FUNCTION_BLOCK ReactorAbortManager (* Basic Function Block Type *)
  (* Standard: 61499-2 *)
  (* Version 0.0, 10/19/2026, Schneider Electric, Template *)
  PACKAGE SE.Nereda;
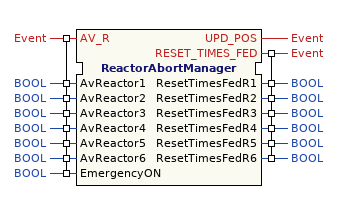
  EVENT_INPUT
    AV_R WITH AvReactor1, AvReactor2, AvReactor3, AvReactor4, AvReactor5, AvReactor6, EmergencyON; (* Normal Execution Request *)
  END_EVENT
  EVENT_OUTPUT
    UPD_POS; (* Execution Confirmation *)
    RESET_TIMES_FED WITH ResetTimesFedR1, ResetTimesFedR2, ResetTimesFedR3, ResetTimesFedR4, ResetTimesFedR5, ResetTimesFedR6;
  END_EVENT
  VAR_INPUT
    AvReactor1 : BOOL;
    AvReactor2 : BOOL;
    AvReactor3 : BOOL;
    AvReactor4 : BOOL;
    AvReactor5 : BOOL;
    AvReactor6 : BOOL;
    EmergencyON : BOOL;
  END_VAR
  VAR_OUTPUT
    ResetTimesFedR1 : BOOL;
    ResetTimesFedR2 : BOOL;
    ResetTimesFedR3 : BOOL;
    ResetTimesFedR4 : BOOL;
    ResetTimesFedR5 : BOOL;
    ResetTimesFedR6 : BOOL;
  END_VAR
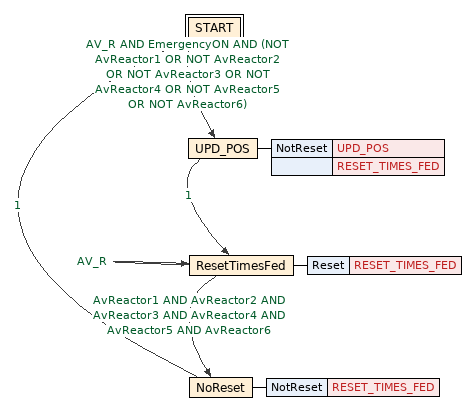
  EC_STATES
    START; (* Initial State *)
    UPD_POS : NotReset -> UPD_POS, -> RESET_TIMES_FED;
    ResetTimesFed : Reset -> RESET_TIMES_FED;
    NoReset : NotReset -> RESET_TIMES_FED;
  END_STATES
  EC_TRANSITIONS
    START TO UPD_POS := AV_R AND EmergencyON AND (NOT AvReactor1 OR NOT AvReactor2 OR NOT AvReactor3 OR NOT AvReactor4 OR NOT AvReactor5 OR NOT AvReactor6);
    UPD_POS TO ResetTimesFed := 1;
    ResetTimesFed TO NoReset := AvReactor1 AND AvReactor2 AND AvReactor3 AND AvReactor4 AND AvReactor5 AND AvReactor6;
    ResetTimesFed TO ResetTimesFed := AV_R;
    NoReset TO START := 1;
  END_TRANSITIONS
  ALGORITHM Reset IN ST:
;
IF NOT AvReactor1 THEN
    ResetTimesFedR1 := TRUE;
END_IF;

IF NOT AvReactor2 THEN
    ResetTimesFedR2 := TRUE;
END_IF;

IF NOT AvReactor3 THEN
    ResetTimesFedR3 := TRUE;
END_IF;

IF NOT AvReactor4 THEN
    ResetTimesFedR4 := TRUE;
END_IF;

IF NOT AvReactor5 THEN
    ResetTimesFedR5 := TRUE;
END_IF;

IF NOT AvReactor6 THEN
	ResetTimesFedR6 := TRUE;
END_IF;
  END_ALGORITHM
  ALGORITHM NotReset IN ST:
;
ResetTimesFedR1 := FALSE;
ResetTimesFedR2 := FALSE;
ResetTimesFedR3 := FALSE;
ResetTimesFedR4 := FALSE;
ResetTimesFedR5 := FALSE;
ResetTimesFedR6 := FALSE;
  END_ALGORITHM
END_FUNCTION_BLOCK
